// TIA Portal project "FactoryIO_Template_S7-1200_V15_V18" (V18)
// Vorlageprojekt für das Buch mit Zielsystem S7-1200

(* hardware
DEVICE "S7-1200-Station_1"  S7-1200 Station
   slot 0: "Baugruppenträger_0"  Rack  V1.0
   slot 1: "PLC_1"  CPU 1214C AC/DC/Rly  6ES7 214-1BG40-0XB0  V4.6
   slot 2: "DQ 16x24VDC_1"  SM 1222 DQ16 x 24VDC  6ES7 222-1BH32-0XB0  V2.0
*)

// ===== PLC "PLC_1"  CPU 1214C AC/DC/Rly =====

VAR_GLOBAL   // PLC tag table "Standard-Variablentabelle"
   "START BUT" AT %I0.0 : Bool;
   "STOP BUT" AT %I0.1 : Bool;
   "RESET BUT" AT %I0.2 : Bool;
   "EMERGENCY BUT" AT %I0.3 : Bool;
   "MAN-AUTO BUT" AT %I0.4 : Bool;
   "SENSOR 1" AT %I0.5 : Bool;
   "SENSOR 2" AT %I0.6 : Bool;
   "SENSOR 3" AT %I0.7 : Bool;
   "URUN TESPIT SENSORU" AT %I1.0 : Bool;
   "KONVEYOR  1" AT %Q0.0 : Bool;
   "KONVEYOR 2" AT %Q0.1 : Bool;
   "TUTUCU" AT %Q0.2 : Bool;
   "X YONUNE GIT" AT %Q0.3 : Bool;
   "Z YONUNE GIT" AT %Q0.4 : Bool;
   "URUN SAYISI" AT %QW8 : Int;
   "START MEM" AT %M10.0 : Bool;
   "URUN TRANSFER MEM" AT %M10.1 : Bool;
   "Tag_1" AT %M10.2 : Bool;
   "SISTEM RESET MEM" AT %M10.3 : Bool;
END_VAR

// folder: System blocks/Program resources

DATA_BLOCK "TIMER 1"   // DB1
{ S7_Optimized_Access := 'TRUE' }
AUTHOR : Simatic
FAMILY : IEC
NAME : IEC_TMR
VERSION : 1.0
// stored: InstanceOfName IEC_TIMER
"IEC_TIMER"
BEGIN
END_DATA_BLOCK

DATA_BLOCK "TIMER 2"   // DB2
{ S7_Optimized_Access := 'TRUE' }
AUTHOR : Simatic
FAMILY : IEC
NAME : IEC_TMR
VERSION : 1.0
// stored: InstanceOfName IEC_TIMER
"IEC_TIMER"
BEGIN
END_DATA_BLOCK

DATA_BLOCK "TIMER 3"   // DB3
{ S7_Optimized_Access := 'TRUE' }
AUTHOR : Simatic
FAMILY : IEC
NAME : IEC_TMR
VERSION : 1.0
// stored: InstanceOfName IEC_TIMER
"IEC_TIMER"
BEGIN
END_DATA_BLOCK

DATA_BLOCK "TIMER 4"   // DB4
{ S7_Optimized_Access := 'TRUE' }
AUTHOR : Simatic
FAMILY : IEC
NAME : IEC_TMR
VERSION : 1.0
// stored: InstanceOfName IEC_TIMER
"IEC_TIMER"
BEGIN
END_DATA_BLOCK

DATA_BLOCK "TIMER 5"   // DB5
{ S7_Optimized_Access := 'TRUE' }
AUTHOR : Simatic
FAMILY : IEC
NAME : IEC_TMR
VERSION : 1.0
// stored: InstanceOfName IEC_TIMER
"IEC_TIMER"
BEGIN
END_DATA_BLOCK

DATA_BLOCK "TIMER 6"   // DB6
{ S7_Optimized_Access := 'TRUE' }
AUTHOR : Simatic
FAMILY : IEC
NAME : IEC_TMR
VERSION : 1.0
// stored: InstanceOfName IEC_TIMER
"IEC_TIMER"
BEGIN
END_DATA_BLOCK

// folder: (top level)

FUNCTION "MHJ-PLC-Lab-Function-S71200" : Void   // FC9000, SCL
{ S7_Optimized_Access := 'TRUE' }
VERSION : 0.1
   VAR_TEMP
      rdTimeReturn : Int;
      outputTime : DTL;
      SyncVal : Byte;
      forVal : Int;
      forVal_2 : Int;
      Value : Byte;
   END_VAR
   VAR CONSTANT
      CompVal : Byte := 16#34;
      Value_01 : Byte := 16#11;
      Value_01_DW : DWord := 16#A165_D992;
      Value_02_DW : DWord := 16#58BE_4401;
   END_VAR
BEGIN

   #Value:=PEEK(area := 16#82,
        dbNumber := 0,
        byteOffset := 511);
   #Value := #Value + 1;

   POKE(area := 16#82,
        dbNumber := 0,
        byteOffset := 511,
        value := #Value);

   POKE(area:=16#81,
        dbNumber:=0,
        byteOffset:=1016,
        value:=#Value_01_DW);
   POKE(area := 16#81,
        dbNumber := 0,
        byteOffset := 1020,
        value := #Value_02_DW);

   POKE(area := 16#81,
        dbNumber := 0,
        byteOffset := 511,
        value := B#16#00);

   FOR #forVal := 0 TO 120 DO
       FOR #forVal_2:=0 TO 10 DO
           #rdTimeReturn:=RD_SYS_T(#outputTime);
           #rdTimeReturn := WR_SYS_T(#outputTime);
           #rdTimeReturn := RD_SYS_T(#outputTime);
           #rdTimeReturn := WR_SYS_T(#outputTime);
       END_FOR;
       #SyncVal:= PEEK(area := 16#81,
                      dbNumber := 0,
                      byteOffset := 511);
       IF #SyncVal = #CompVal THEN
          GOTO M_1;
       END_IF;
   END_FOR;
   RETURN;

   M_1:
   POKE(area := 16#81,
        dbNumber := 0,
        byteOffset := 511,
        value := B#16#0);
END_FUNCTION

ORGANIZATION_BLOCK "Main"   // OB1, LAD, ProgramCycle
TITLE = "Main Program Sweep (Cycle)"
{ S7_Optimized_Access := 'TRUE' }
VERSION : 0.1
   VAR_INPUT
      Initial_Call : Bool;   // Initial call of this OB
      Remanence : Bool;   // =True, if remanent data are available
   END_VAR
   VAR_TEMP   // added for the SCL form of the ladder/FBD networks
      _w1 : Bool;
   END_VAR
BEGIN

REGION Network 1: Konnektierungsbaustein für PLC-Lab
   // Im Netzwerk 1 wird der Konnektierungsbaustein für PLC-Lab aufgerufen.
   // Dieser Aufruf darf nicht entfernt werden!
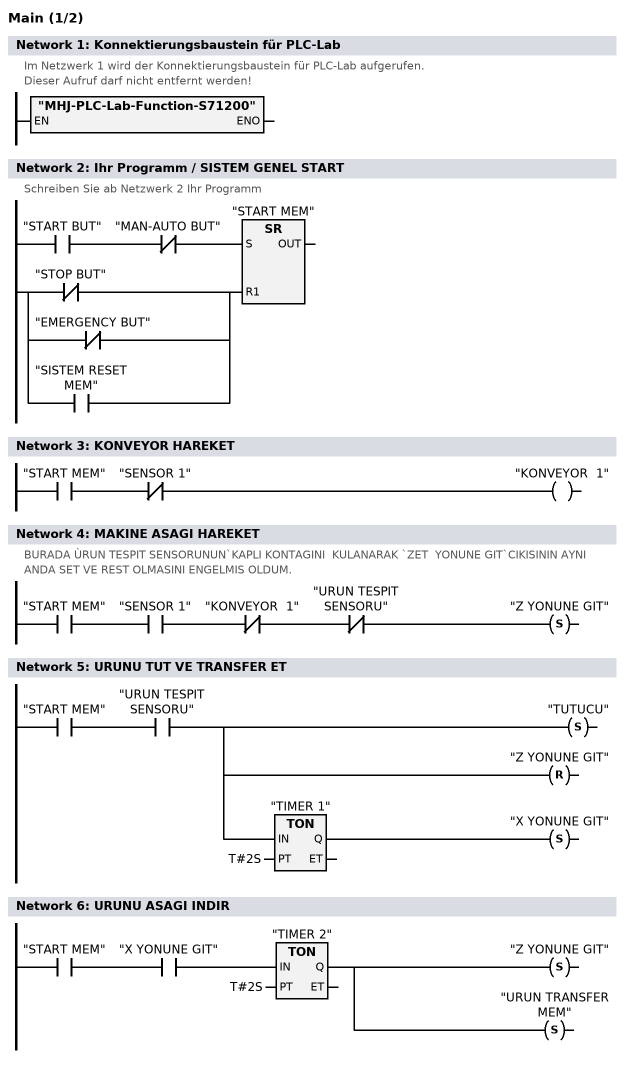
   RUNG wire#powerrail
      "MHJ-PLC-Lab-Function-S71200"()
   END_RUNG
   // the same network as SCL:
   "MHJ-PLC-Lab-Function-S71200"();
END_REGION

REGION Network 2: Ihr Programm / SISTEM GENEL START
   // Schreiben Sie ab Netzwerk 2 Ihr Programm
   RUNG wire#powerrail
      Contact( "START BUT" )
      I_Contact( "MAN-AUTO BUT" )
      S_SR(operand := "START MEM", r1 := wire#w1)
   END_RUNG
   RUNG wire#powerrail
      I_Contact( "STOP BUT" )
   END_RUNG wire#w1
   RUNG wire#powerrail
      I_Contact( "EMERGENCY BUT" )
   END_RUNG wire#w1
   RUNG wire#powerrail
      Contact( "SISTEM RESET MEM" )
   END_RUNG wire#w1
   // the same network as SCL:
   IF "START BUT" AND NOT "MAN-AUTO BUT" THEN
       "START MEM" := TRUE;   // SR flip-flop
   END_IF;
   IF NOT "STOP BUT" OR NOT "EMERGENCY BUT" OR "SISTEM RESET MEM" THEN "START MEM" := FALSE; END_IF;
END_REGION

REGION Network 3: KONVEYOR HAREKET
   RUNG wire#powerrail
      Contact( "START MEM" )
      I_Contact( "SENSOR 1" )
      Coil( "KONVEYOR  1" )
   END_RUNG
   // the same network as SCL:
   "KONVEYOR  1" := "START MEM" AND NOT "SENSOR 1";
END_REGION

REGION Network 4: MAKINE ASAGI HAREKET
   // BURADA ÙRUN TESPIT SENSORUNUN`KAPLI KONTAGINI  KULANARAK `ZET  YONUNE GIT`CIKISININ AYNI ANDA SET VE REST OLMASINI ENGELMIS OLDUM.
   RUNG wire#powerrail
      Contact( "START MEM" )
      Contact( "SENSOR 1" )
      I_Contact( "KONVEYOR  1" )
      I_Contact( "URUN TESPIT SENSORU" )
      S_Coil( "Z YONUNE GIT" )
   END_RUNG
   // the same network as SCL:
   IF "START MEM" AND "SENSOR 1" AND NOT "KONVEYOR  1" AND NOT "URUN TESPIT SENSORU" THEN
       "Z YONUNE GIT" := TRUE;
   END_IF;
END_REGION

REGION Network 5: URUNU TUT VE TRANSFER ET
   #_w1 := "START MEM" AND "URUN TESPIT SENSORU";
   IF #_w1 THEN
       "TUTUCU" := TRUE;
       "Z YONUNE GIT" := FALSE;
   END_IF;
   "TIMER 1".TON(IN := #_w1, PT := T#2S);
   IF "TIMER 1".Q THEN "X YONUNE GIT" := TRUE; END_IF;
END_REGION

REGION Network 6: URUNU ASAGI INDIR
   "TIMER 2".TON(IN := "START MEM" AND "X YONUNE GIT", PT := T#2S);
   IF "TIMER 2".Q THEN
       "Z YONUNE GIT" := TRUE;
       "URUN TRANSFER MEM" := TRUE;
   END_IF;
END_REGION

REGION Network 7: URUNU BIRAK VE ILK KONUMUNA DON
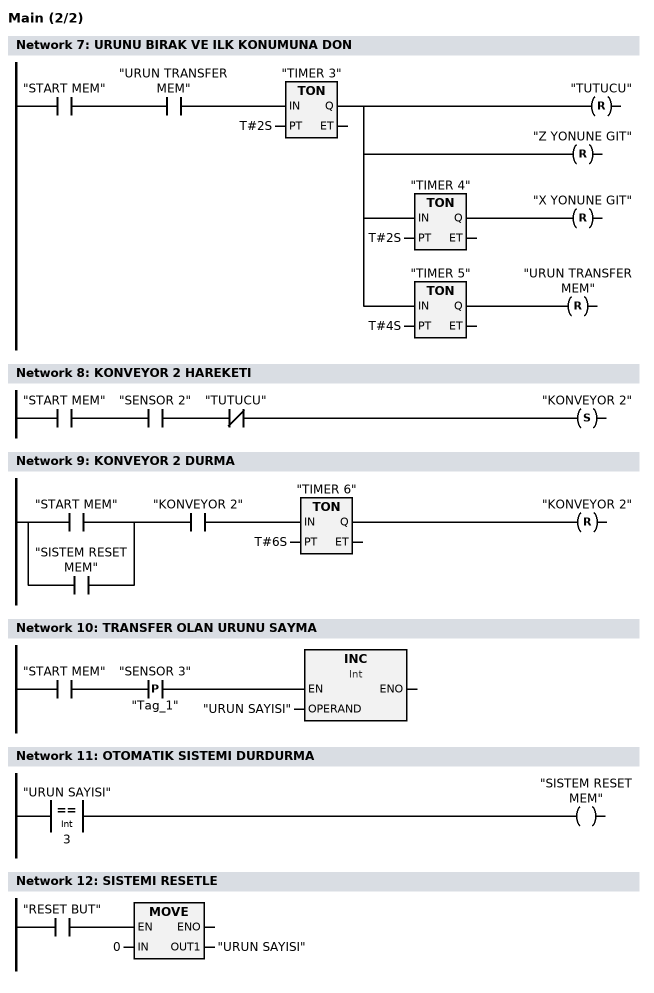
   "TIMER 3".TON(IN := "START MEM" AND "URUN TRANSFER MEM", PT := T#2S);
   IF "TIMER 3".Q THEN
       "TUTUCU" := FALSE;
       "Z YONUNE GIT" := FALSE;
   END_IF;
   "TIMER 4".TON(IN := "TIMER 3".Q, PT := T#2S);
   IF "TIMER 4".Q THEN "X YONUNE GIT" := FALSE; END_IF;
   "TIMER 5".TON(IN := "TIMER 3".Q, PT := T#4S);
   IF "TIMER 5".Q THEN "URUN TRANSFER MEM" := FALSE; END_IF;
END_REGION

REGION Network 8: KONVEYOR 2 HAREKETI
   RUNG wire#powerrail
      Contact( "START MEM" )
      Contact( "SENSOR 2" )
      I_Contact( "TUTUCU" )
      S_Coil( "KONVEYOR 2" )
   END_RUNG
   // the same network as SCL:
   IF "START MEM" AND "SENSOR 2" AND NOT "TUTUCU" THEN "KONVEYOR 2" := TRUE; END_IF;
END_REGION

REGION Network 9: KONVEYOR 2 DURMA
   "TIMER 6".TON(IN := ("START MEM" OR "SISTEM RESET MEM") AND "KONVEYOR 2", PT := T#6S);
   IF "TIMER 6".Q THEN "KONVEYOR 2" := FALSE; END_IF;
END_REGION

REGION Network 10: TRANSFER OLAN URUNU SAYMA
   RUNG wire#powerrail
      Contact( "START MEM" )
      P_Contact(operand := "SENSOR 3", bit := "Tag_1")
      { S7_Templates := "DestType := Int" } Inc( "URUN SAYISI" )
   END_RUNG
   // the same network as SCL:
   #_w1 := "START MEM" AND "SENSOR 3" AND NOT "Tag_1";   // rising edge of "SENSOR 3"
   "Tag_1" := "SENSOR 3";
   IF #_w1 THEN "URUN SAYISI" := "URUN SAYISI" + 1; END_IF;
END_REGION

REGION Network 11: OTOMATIK SISTEMI DURDURMA
   RUNG wire#powerrail
      { S7_Templates := "SrcType := Int" } EQ_Contact(in1 := "URUN SAYISI", in2 := 3)
      Coil( "SISTEM RESET MEM" )
   END_RUNG
   // the same network as SCL:
   "SISTEM RESET MEM" := "URUN SAYISI" = 3;
END_REGION

REGION Network 12: SISTEMI RESETLE
   RUNG wire#powerrail
      Contact( "RESET BUT" )
      Move(in := 0, out1 => "URUN SAYISI")
   END_RUNG
   // the same network as SCL:
   IF "RESET BUT" THEN "URUN SAYISI" := 0; END_IF;
END_REGION
END_ORGANIZATION_BLOCK